// TIA Portal V21 export
// export: Created 2026-11-21T23:19:45.2483508Z, ExportSetting WithDefaults, DisplayName Totally Integrated Automation Portal, DisplayVersion V21 Update 3, DisplayName STEP 7 Professional, DisplayVersion V21 Update 3, DisplayName STEP 7 Safety, DisplayVersion V21, DisplayName Tech WebApplication, DisplayVersion V21, DisplayName WinCC Basic/Comfort/Advanced, DisplayVersion V21 Update 3, DisplayName WinCC Unified, DisplayVersion V21 Update 3
Screen "Ctl_03_UserView"  1024x768, Number=12, Template=Nav
  ScreenLayer 
    UserView "User view_1" at 3,3 size 480x240  Appearance=AppearanceFlat, CountVisibleItems=8, ViewType=ViewTypeComplex
